// TIA Portal V21 export
FUNCTION_BLOCK "FB_Sequence"   // FB21, GRAPH
BEGIN
END_FUNCTION_BLOCK
